Fanuc KAREL source: KC00043.KL

PROGRAM KC00043
%NOLOCKGROUP
%ENVIRONMENT REGOPE
VAR
  I: INTEGER
  J: INTEGER
  K: INTEGER
  R: REAL
  B: BOOLEAN
  S: STRING[80]
  T: STRING[80]
  P: PATH
  Q: PATH
  AI: ARRAY[8] OF INTEGER
  AB: ARRAY[244] OF BYTE
  EP: XYZWPREXT
BEGIN
  EP = GET_TPE_POS_REG(I,J)
END KC00043
